ABB RAPID module: LongProg_0.mod

%%%
  VERSION:1
  LANGUAGE:ENGLISH
%%%
MODULE MOD_Tmp1

	PROC Prg_Tmp1()

		ConfJ \On;
		ConfL \Off;
		! Program generated by RoboDK v6.0.7 for ABB IRBT 2005 Standard 2.8m on XX/XX/XXXX 18:00:00
		! Using nominal kinematics.
		MoveAbsJ [[250.000000,0.000000,0.000000,0.000000,0.000000,0.000000],[9E+09,9E+09,9E+09,9E+09,9E+09,9E+09]],v500,z1,ToolS \WObj:=FrameS;

	ENDPROC

ENDMODULE
